// TIA Portal V20 export
// export: Created 2026-10-12T04:58:20.1136826Z, ExportSetting WithDefaults, DisplayName Totally Integrated Automation Portal, DisplayVersion V20, DisplayName TIA Portal Openness, DisplayVersion V20, DisplayName TIA Portal Teamcenter Gateway, DisplayVersion V20, DisplayName TIA Portal Version Control Interface, DisplayVersion V20, DisplayName SINAMICS Startdrive Advanced, DisplayVersion V20 SP1 Update 2, DisplayName SINAMICS Startdrive G110M, G120, G120C, G120D, G120P, G115D, DisplayVersion V20 SP1 Update 2, DisplayName SINAMICS Startdrive G130, G150, S120, S150, SINAMICS MV, G220, S200, S210, DisplayVersion V20 SP1 Update 2, DisplayName STEP 7 Professional, DisplayVersion V20, DisplayName STEP 7 Safety, DisplayVersion V20, DisplayName WinCC Basic/Comfort/Advanced, DisplayVersion V20, DisplayName WinCC Professional, DisplayVersion V20, DisplayName WinCC Unified, DisplayVersion V20
FUNCTION "FRK_AccessPolicyCrc" : DWord   // FC56, SCL
{ S7_Optimized_Access := 'TRUE' }
VERSION : 0.1
// stored: AutoNumber true, IsIECCheckEnabled false, SetENOAutomatically false, UDAEnableTagReadback false
   VAR_IN_OUT
      Image : "FRK_AccessPolicyImage";
   END_VAR
   VAR_TEMP
      Work : DWord;
      Index : Int;
      Size : Int;
   END_VAR
BEGIN

   #Work := "FRK_AccessCrcNumber"(Previous := DWORD#16#FFFFFFFF, Value := UINT_TO_UDINT(#Image.SchemaVersion));
   #Work := "FRK_AccessCrcNumber"(Previous := #Work, Value := #Image.Generation);
   #Size := LEN(#Image.Scope);
   #Work := "FRK_AccessCrcNumber"(Previous := #Work, Value := INT_TO_UDINT(#Size));
   FOR #Index := 1 TO #Size DO
       #Work := "FRK_AccessCrcByte"(Previous := #Work, Value := CHAR_TO_BYTE(#Image.Scope[#Index]));
   END_FOR;
   FOR #Index := 0 TO 11 DO
       #Work := "FRK_AccessCrcNumber"(Previous := #Work, Value := DINT_TO_UDINT(#Image.Policy.Required[#Index]));
   END_FOR;
   #Work := "FRK_AccessCrcNumber"(Previous := #Work, Value := DINT_TO_UDINT(TIME_TO_DINT(#Image.Policy.SessionTimeout)));
   #FRK_AccessPolicyCrc := NOT #Work;
END_FUNCTION
